Fanuc KAREL source: kt00743.KL

-- PROVISIONAL review KL for V1013-1; original PC SHA256 d0992907ebbc2c80d62978bf06d6f053fa165dec0e4714c08473edf39192bd17
-- Incomplete behavior may be omitted. Consult companion uncertainty JSON. Do not deploy.
PROGRAM KT00743
%NOLOCKGROUP
VAR
  OUT : INTEGER
-- UNRESOLVED_DECL ARG type=002013
BEGIN
  -- UNRESOLVED_PC offsets 5-18; opcodes 22,1D,23
  -- UNRESOLVED_PC offsets 23-27; opcodes 7F
END KT00743
